Fanuc KAREL source: kc00012.KL

-- PROVISIONAL review KL for V770-1; original PC SHA256 0803982cf17807eea4bfe9d4acc3ba904b52dd63d92211a44078cfbd1f45a123
-- Incomplete behavior may be omitted. Consult companion uncertainty JSON. Do not deploy.
PROGRAM KC00012
%NOLOCKGROUP
BEGIN
  -- UNRESOLVED_PC offsets 5-51; opcodes 27,22,22,22,22,22,22,22,31
  -- UNRESOLVED_PC offsets 56-60; opcodes 7F
END KC00012
